Fanuc KAREL source: kc00016.KL

-- PROVISIONAL review KL for V1013-1; original PC SHA256 e758a18466d8b73d9aa3022a95fb7fe723f209eae393856a0122aec1d7c2a1da
-- Incomplete behavior may be omitted. Consult companion uncertainty JSON. Do not deploy.
PROGRAM KC00016
%NOLOCKGROUP
BEGIN
  -- UNRESOLVED_PC offsets 5-15; opcodes 27,22,31
  -- UNRESOLVED_PC offsets 20-24; opcodes 7F
END KC00016
